(* IEC 61131-3 sources: sceptre-phenix-topologies/cherrymountain-brewery/plant/generated/lite/openplc/plc-brewhouse, 1 file *)

(* ---- located_vars.st ---- *)
(* Generated by plantgen from plant/plant.yaml (variant lite). Do not edit. *)
(* Analog values are raw registers: engineering value = raw / 10^scaling. *)
(* RIO I/O is at %IX100.0 / %QX100.0 / %IW100 / %QW100 (v3 and v4 alike). *)
(* PLC memory: bits from %QX0.0 (coils), words from %MW0 (holding register qw_count and up, see modbus_slave.json). *)
VAR
  BH_MILL_LT01_PV AT %IW100 : UINT; (* Grain silo level, %, x10 *)
  BH_MILL_SI01_PV AT %IW101 : UINT; (* Mill VFD speed, Hz, x10 *)
  BH_MILL_YS01_PV AT %IX100.0 : BOOL; (* Mill running *)
  BH_MILL_HS01_CMD AT %QX100.0 : BOOL; (* Mill run command *)
  BH_MILL_HS02_CMD AT %QX100.1 : BOOL; (* Grain auger run command *)
  BH_MILL_SC01_SP AT %QW100 : UINT; (* Mill VFD speed reference, Hz, x10 *)
  BH_CLT_LT01_PV AT %IW102 : UINT; (* CLT level, %, x10 *)
  BH_CLT_TT01_PV AT %IW103 : UINT; (* CLT temperature, degF, x10 *)
  BH_CLT_LSH01_PV AT %IX100.1 : BOOL; (* CLT high-level switch *)
  BH_CLT_XV01_CMD AT %QX100.2 : BOOL; (* CLT fill valve (RO permeate) *)
  BH_HLT_LT01_PV AT %IW104 : UINT; (* HLT level, %, x10 *)
  BH_HLT_LT01_ALM_LOW AT %QX0.0 : BOOL; (* HLT level: low alarm (low) *)
  BH_HLT_TT01_PV AT %IW105 : UINT; (* HLT temperature, degF, x10 *)
  BH_HLT_TT01_ALM_HIGH AT %QX0.1 : BOOL; (* HLT temperature: high alarm (medium) *)
  BH_HLT_LSL01_PV AT %IX100.2 : BOOL; (* HLT low-level switch (made while the steam jacket is covered; drops below 15 %) *)
  BH_HLT_XV01_CMD AT %QX100.3 : BOOL; (* HLT fill valve (from the CLT) *)
  BH_HLT_TV01_OUT AT %QW101 : UINT; (* HLT steam valve position, %, x10 *)
  BH_HLT_TT01_SP AT %MW0 : UINT; (* HLT temperature setpoint, degF, x10 *)
  BH_MLT_TT01_PV AT %IW106 : UINT; (* MLT mash temperature, degF, x10 *)
  BH_MLT_TT01_ALM_DEVIATION AT %QX0.2 : BOOL; (* MLT mash temperature: deviation alarm (medium) *)
  BH_MLT_LT01_PV AT %IW107 : UINT; (* MLT level, %, x10 *)
  BH_MLT_PDT01_PV AT %IW108 : UINT; (* MLT false-bottom differential pressure, psi, x100 *)
  BH_MLT_PDT01_ALM_HIGH AT %QX0.3 : BOOL; (* MLT false-bottom differential pressure: high alarm (medium) *)
  BH_MLT_FT01_PV AT %IW109 : UINT; (* Lauter runoff flow, gal/min, x10 *)
  BH_MLT_FT02_PV AT %IW110 : UINT; (* Sparge flow, gal/min, x10 *)
  BH_MLT_ZT01_PV AT %IW111 : UINT; (* Rake height above the false bottom, in, x10 *)
  BH_MLT_YS01_PV AT %IX100.3 : BOOL; (* Rake running *)
  BH_MLT_XV01_CMD AT %QX100.4 : BOOL; (* Strike water valve (from the HLT) *)
  BH_MLT_HS01_CMD AT %QX100.5 : BOOL; (* Rake run command *)
  BH_MLT_TV01_OUT AT %QW102 : UINT; (* MLT jacket steam valve position, %, x10 *)
  BH_MLT_FV01_OUT AT %QW103 : UINT; (* Runoff valve position, %, x10 *)
  BH_MLT_FV02_OUT AT %QW104 : UINT; (* Sparge valve position, %, x10 *)
  BH_MLT_SC01_OUT AT %QW105 : UINT; (* Rake speed reference, %, x10 *)
  BH_MLT_TT01_SP AT %MW1 : UINT; (* Mash step temperature setpoint, degF, x10 *)
  BH_MLT_XS01_ACTIVE AT %QX0.4 : BOOL; (* Mash step at temperature, or 15 min into it (deviation alarm enabled) *)
  BH_KTL_TT01_PV AT %IW112 : UINT; (* Kettle temperature, degF, x10 *)
  BH_KTL_LT01_PV AT %IW113 : UINT; (* Kettle level, %, x10 *)
  BH_KTL_LT01_ALM_HIGH AT %QX0.5 : BOOL; (* Kettle level: high alarm (high) *)
  BH_KTL_PT01_PV AT %IW114 : UINT; (* Ambient (barometric) pressure for boil detection, psia, x100 *)
  BH_KTL_LSH01_PV AT %IX100.4 : BOOL; (* Kettle high-level switch (boil-over) *)
  BH_KTL_XV01_CMD AT %QX100.6 : BOOL; (* Whirlpool tangential inlet valve *)
  BH_KTL_XV02_CMD AT %QX100.7 : BOOL; (* Whirlpool hop doser *)
  BH_KTL_TV01_OUT AT %QW106 : UINT; (* Kettle jacket steam valve position, %, x10 *)
  BH_KTL_TB01_PV AT %MW2 : UINT; (* Computed local wort boiling point, degF, x10 *)
  BH_KTL_KI01_PV AT %MW3 : UINT; (* Boil time elapsed, min, x10 *)
  BH_KTL_XS01_BOIL AT %QX0.6 : BOOL; (* Boil detected (within 0.5 degF of the boiling point) *)
  BH_KO_FT01_PV AT %IW115 : UINT; (* Wort flow to the fermenter, gal/min, x10 *)
  BH_KO_TT01_PV AT %IW116 : UINT; (* HX stage-1 wort outlet temperature (CLT water side), degF, x10 *)
  BH_KO_TT02_PV AT %IW117 : UINT; (* Knockout wort temperature (after stage 2), degF, x10 *)
  BH_KO_TT02_ALM_DEVIATION AT %QX0.7 : BOOL; (* Knockout wort temperature (after stage 2): deviation alarm (high) *)
  BH_KO_FT02_PV AT %IW118 : UINT; (* Inline O2 flow, L/min, x100 *)
  BH_KO_AT01_PV AT %IW119 : UINT; (* Wort dissolved oxygen, ppm, x100 *)
  BH_KO_AT01_ALM_LOW AT %QX1.0 : BOOL; (* Wort dissolved oxygen: low alarm (low) *)
  BH_KO_YS01_PV AT %IX100.5 : BOOL; (* Wort pump running *)
  BH_KO_HS01_CMD AT %QX101.0 : BOOL; (* Wort pump run command *)
  BH_KO_XV01_CMD AT %QX101.1 : BOOL; (* Knockout valve to the fermenter header *)
  BH_KO_SC01_OUT AT %QW107 : UINT; (* Wort pump VFD speed reference, %, x10 *)
  BH_KO_TV01_OUT AT %QW108 : UINT; (* HX stage-2 glycol valve position, %, x10 *)
  BH_KO_FC01_SP AT %QW109 : UINT; (* Inline O2 mass-flow setpoint, L/min, x100 *)
  BH_KO_TT02_SP AT %MW4 : UINT; (* Knockout temperature setpoint, degF, x10 *)
  BH_BATCH_XC01_PHASE AT %MW5 : UINT; (* Phase selected by the batch engine, None, x1 *)
  BH_BATCH_XC01_CMD AT %MW6 : UINT; (* Phase command, None, x1 *)
  BH_BATCH_XS01_STATE AT %MW7 : UINT; (* Phase state, None, x1 *)
  BH_BATCH_XS01_STEP AT %MW8 : UINT; (* Phase step number, None, x1 *)
  BH_BATCH_XI01_BATCH AT %MW9 : UINT; (* Batch number (low 16 bits), None, x1 *)
  BH_BATCH_XC03_PARAM AT %MW10 : UINT; (* Phase parameter (MILL kg, MASH_IN liters, MASH_STEP, BOIL, and WHIRLPOOL minutes; 0 = program default), None, x1 *)
  BH_BATCH_XI02_REQUESTS AT %IW120 : UINT; (* Brews requested at the brewhouse panel since the start (16-bit counter), None, x1 *)
  BH_BATCH_XC02_ACCEPTED AT %MW11 : UINT; (* Brew requests the batch engine has accepted (16-bit counter; the engine writes it), None, x1 *)
  BH_BATCH_XI03_ACCEPTED AT %QW110 : UINT; (* Accepted-request counter sent to the panel (the program forwards XC02), None, x1 *)
  BH_ENTRY_HS01_ENTRY AT %QX1.1 : BOOL; (* MLT entry permit issued (entry supervisor; locks the vessel out) *)
  BH_ENTRY_HS02_ENTRY AT %QX1.2 : BOOL; (* Kettle entry permit issued (entry supervisor; locks the vessel out) *)
  BH_ENTRY_XS01_LOCKED AT %QX1.3 : BOOL; (* MLT locked out for entry (steam, strike and sparge water, runoff, rake) *)
  BH_ENTRY_XS02_LOCKED AT %QX1.4 : BOOL; (* Kettle locked out for entry (steam, whirlpool, hop doser) *)
  BH_ENTRY_XA01_PV AT %QX1.5 : BOOL; (* MLT write or phase start against a locked-out output during entry *)
  BH_ENTRY_XA01_ALM_STATE AT %QX1.6 : BOOL; (* MLT write or phase start against a locked-out output during entry: state alarm (critical) *)
  BH_ENTRY_XA02_PV AT %QX1.7 : BOOL; (* Kettle write or phase start against a locked-out output during entry *)
  BH_ENTRY_XA02_ALM_STATE AT %QX2.0 : BOOL; (* Kettle write or phase start against a locked-out output during entry: state alarm (critical) *)
END_VAR
